(* IEC 61131-3 sources: rusty/tests/lit/cfc/generics/generic_output, 2 files *)

(* ---- main.st ---- *)
FUNCTION main : DINT
    generic_output.x := 21;
    generic_output();
    // CHECK: y = 42
    printf('y = %d$N', generic_output.y);
END_FUNCTION

(* ---- myGenOut.st ---- *)
FUNCTION myGenOut<T: ANY_NUM>
VAR_INPUT
    a : T;
END_VAR
VAR_OUTPUT
    doubled : T;
END_VAR
END_FUNCTION

FUNCTION myGenOut__DINT
VAR_INPUT
    a : DINT;
END_VAR
VAR_OUTPUT
    doubled : DINT;
END_VAR
    doubled := a * 2;
END_FUNCTION
